(* IEC 61131-3 sources: Elmo_Master/Lasal_PRG/MotionTCPDemo/Class/ReceiveMsg, 1 file *)

(* ---- ReceiveMsg.st ---- *)
(*!
<Class
	Name               = "ReceiveMsg"
	Revision           = "0.0"
	RealtimeTask       = "false"
	CyclicTask         = "false"
	BackgroundTask     = "true"
	Sigmatek           = "false"
	OSInterface        = "false"
	HighPriority       = "false"
	Automatic          = "false"
	UpdateMode         = "Prescan"
	SharedCommandTable = "true"
	Objectsize         = "(284,120)">
	<Channels>
		<Server Name="Msg" Visualized="false" Initialize="false" WriteProtected="true" Retentive="false"/>
	</Channels>
	<Network Name="ReceiveMsg">
		<!-- List of Components in this network -->
		<Components>
			<Object
				Name       = "_base"
				Class      = "_SigTCPComReceive"
				Position   = "(218,120)"
				Visualized = "false">
				<Channels>
					<Server Name="ClassSvr"/>
					<Server Name="RecvCnt"/>
					<Server Name="SourceID"/>
					<Client Name="_SigTCPDataManager"/>
				</Channels>
			</Object>
		</Components>
		<Comments>
		</Comments>
		<!-- List of Connections in this network -->
		<Connections>
			<Connection Source="this.ClassSvr" Destination="_base.ClassSvr" Vertices="(1006,210),(834,210),"/>
			<Connection Source="this.SourceID" Destination="_base.SourceID" Vertices="(1006,270),(834,270),"/>
			<Connection Source="this.RecvCnt" Destination="_base.RecvCnt" Vertices="(1006,330),(834,330),"/>
			<Connection Source="_base._SigTCPDataManager" Destination="this._SigTCPDataManager" Vertices="(218,210),(38,210),"/>
		</Connections>
		<!-- Headerfiles -->
		<Options>
		</Options>
	</Network>
</Class>
*)
#pragma using _SigTCPComReceive

ReceiveMsg : CLASS
: _SigTCPComReceive
  //Servers:
	Msg 	: SvrCh_DINT;
  //Clients:
  //Variables:
  //Functions:
				//! <Function Comment="Is called whenever data is received. &#13;&#10;Overwrite this method to process data. &#13;&#10;NOTE: If the optional CMD parameter is used when sending, the method CallBackReciverCMD() has to be used for receiving in order to correctly receive the CMD parameter." Name="CallBackReceiver"/>
	FUNCTION VIRTUAL GLOBAL CallBackReceiver
		VAR_INPUT
			DestinationID 	: DINT;			//! <Variable Comment="ID of Destination.&#13;&#10;ID like in the send object of the remote station in DestinationID." Name="CallBackReceiver.DestinationID"/>
			SourceID 	: DINT;			//! <Variable Comment="ID of Source.&#13;&#10;ID like in the send object of the remote station in SourceID." Name="CallBackReceiver.SourceID"/>
			size 	: UDINT;			//! <Variable Comment="Length of the data received in bytes" Name="CallBackReceiver.size"/>
			pdata 	: ^USINT;			//! <Variable Comment="Pointer to received data" Name="CallBackReceiver.pdata"/>
		END_VAR
		VAR_OUTPUT
			retcode 	: BOOL;			//! <Variable Comment="TRUE = successfully received = _MNG_Recived &#13;&#10;FALSE = Error in receiving = _MNG_GlobalReciveError&#13;&#10;&#13;&#10;Here you can influence how to react on received data packets. &#13;&#10;If FALSE is returned here, an error is triggered in the sending station (see CallbackJobState in the documentation of the class _SigTCPComSend). " Name="CallBackReceiver.retcode"/>
		END_VAR;
  //Tables:
	FUNCTION @STD
		VAR_OUTPUT
			ret_code	: CONFSTATES;
		END_VAR;
	FUNCTION GLOBAL TAB @CT_;
END_CLASS;

FUNCTION VIRTUAL GLOBAL ReceiveMsg::CallBackReceiver
	VAR_INPUT
		DestinationID 	: DINT;
		SourceID 	: DINT;
		size 	: UDINT;
		pdata 	: ^USINT;
	END_VAR
	VAR_OUTPUT
		retcode 	: BOOL;
	END_VAR

  Msg := pdata^$DINT;

END_FUNCTION
